TYPE "ST_DecisionRequest"
VERSION : 0.1
   STRUCT
      "Prompt" : WString[255];
      "Options" : Array[1..6] of String[64];
      "Default" : Int;
      "Timeout" : Time;
      "SourcePath" : WString[255];
   END_STRUCT;
END_TYPE
